Fanuc KAREL source: ks00018.KL

PROGRAM KS00018
%STACKSIZE=65535
%PRIORITY=65535
%NOLOCKGROUP
VAR
A : FILE
B : FILE
FLAG : BOOLEAN
N : INTEGER
STATUS : INTEGER
PN : STRING[80]
VN : STRING[80]
BEGIN
PN=''
VN='A'
-- UNRESOLVED_PC line 19 opcodes [22 63 23] marker_code=27
END KS00018
